{attribute 'qualified_only'}
VAR_GLOBAL RETAIN
	ShutterR1Config : stShutterConfig :=(HeightTravelTime := T#15S,
										HeightTravelTimeOverstep := T#1S,
										AngleTravelTime := T#2S);
END_VAR

(* stored: Version 1.1.0.1
   GVL gvlShutters: Id {14207c95-03ef-4fbc-b845-1f2852642cd2} *)
